(* PLC project zarechnaya.project, CODESYS CODESYS V3.5 SP17 Patch 3 *)
(* stored: creationDateTime 2026-10-20T05:42:22.312171, modificationDateTime 1601-01-01T03:00:00 *)

(* PRG_FilterAlt — выбор режима фильтрации (SFC, PROGRAM: альтернатива, прыжок, приоритет переходов). Шаги: Wait (начальный) → альтернатива слева направо: [xHigh] → Fast, [xLow] → Slow (оба TRUE — побеждает левый, Fast); Fast → [NOT xHigh] и Slow → [NOT xLow] → Done → [xReset] сходятся и прыжком возвращаются на Wait. (Ветви, оканчивающиеся прыжком без схождения, CODESYS 3.5.17 из PLCopen молча не импортирует — проверено на этом кейсе 20.10.2026.) Действия (IEC, N): Fast — ActFast (iFast += 1), Slow — ActSlow (iSlow += 1), Done — ActDone (iDone += 1). *)
PROGRAM PRG_FilterAlt
  VAR_INPUT
    xHigh : BOOL;
    xLow : BOOL;
    xReset : BOOL;
  END_VAR
  VAR_OUTPUT
    iFast : INT;
    iSlow : INT;
    iDone : INT;
  END_VAR

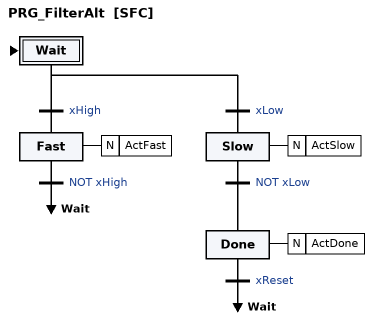
INITIAL_STEP Wait:
END_STEP
TRANSITION FROM Wait TO Fast
  := xHigh;
END_TRANSITION
TRANSITION FROM Wait TO Slow
  := xLow;
END_TRANSITION
STEP Fast:
  ActFast(N);
END_STEP
TRANSITION FROM Fast TO Wait
  := NOT xHigh;
END_TRANSITION
STEP Slow:
  ActSlow(N);
END_STEP
TRANSITION FROM Slow TO Done
  := NOT xLow;
END_TRANSITION
STEP Done:
  ActDone(N);
END_STEP
TRANSITION FROM Done TO Wait
  := xReset;
END_TRANSITION

ACTION ActFast:
                iFast := iFast + 1;

              
END_ACTION

ACTION ActSlow:
                iSlow := iSlow + 1;

              
END_ACTION

ACTION ActDone:
                iDone := iDone + 1;

              
END_ACTION
END_PROGRAM
